(* IEC 61131-3 sources: Codesys_IAP/Demo/PLC1/Magazijn Overzetter Simulatie Structured Text 2V1_tekst/Simulatie, 5 files *)

(* ---- MagazijnDUT.st ---- *)
(*#### DECLARATIE ####*)
{attribute 'qualified_only'}
{attribute 'strict'}
TYPE MagazijnDUT :
(
	INGETROKKEN, INTREKKEN, UITGESTOTEN, UITSTOTEN, LEEG
);
END_TYPE

(* ---- OverzetterDUT.st ---- *)
(*#### DECLARATIE ####*)
{attribute 'qualified_only'}
{attribute 'strict'}
TYPE OverzetterDUT :
(
	INHETMIDDEN, NAARRECHTS, ISRECHTS, NAARLINKS, ISLINKS, GEVALLEN
);
END_TYPE

(* ---- SIM.st ---- *)
(*#### DECLARATIE ####*)
{attribute 'qualified_only'}
VAR_GLOBAL
	// Rotatie van de overzetter
	Vx_OvzRotate: INT := 0;
	// Visualisatie invisible blok
	Vx_OvzBlokLinks: BOOL := FALSE;
	// Visualisatie invisible blok
	Vx_OvzBlokOverzetter: BOOL := FALSE;
	// Visualisatie invisible blok
	Vx_OvzBlokRechts: BOOL := FALSE;
	// Visualisatie invisible blok
	Vx_OvzBlokGevallen: BOOL := FALSE;
	// Magazijn opnieuw vullen (simulatie)
	Ix_MagazijnVullen 	: BOOL;
	// Simulatie visualisatie
	Vw_Rotate45: INT := 45;
	// Visualisatie X positie van de uitstoter
	Vw_MagUitstoterBekerX: INT := 30;
	// Visualisatie invisible blok uitgestoten
	Vx_MagBlokUit: BOOL := TRUE;
	// Visualisatie invisible blok 1
	Vx_MagBlok1: BOOL := TRUE;
	// Visualisatie invisible blok 2
	Vx_MagBlok2: BOOL := TRUE;
	// Visualisatie invisible blok 3
	Vx_MagBlok3: BOOL := TRUE;
	// Visualisatie invisible blok 4
	Vx_MagBlok4: BOOL := TRUE;
	// Visualisatie invisible blokken
	Vx_MagBlok: ARRAY[1..8] OF BOOL;
	// Aantal blokken in het magazijn
	Vw_MagBlokAantal: INT := 4;
	// Simulatie onthoudt dat een blok maar 1x wordt uitgestoten
	Vw_MagBlok1X: INT := 0;
	// Simulatie error. Inverse logica.
	Vx_MagLuchtDrukError: BOOL := TRUE;
	// Simulatie error. Inverse logica.
	Vx_MagIsInError: BOOL := TRUE;
	// Simulatie error. Inverse logica.
	Vx_MagIsUitError: BOOL := TRUE;
	// Simulatie error. Inverse logica.
	Vx_OvzLuchtDrukError: BOOL := TRUE;
	// Simulatie error. Inverse logica.
	Vx_OvzIsLinksError: BOOL := TRUE;
	// Simulatie error. Inverse logica.
	Vx_OvzIsRechtsError: BOOL := TRUE;
	// Simulatie error. Inverse logica.
	Vx_OvzVacuumError: BOOL := TRUE;
	// Kleur van de blokken in het magazijn (lege plek = grijs)
	Vw_MagKleur: ARRAY[1..8] OF DWORD;
	// Kleur van het uitgestoten blok
	Vw_MagKleurUit: DWORD;
	// Kleur van het blok op de overzetter
	Vw_OvzKleur: DWORD := 16#FFC0C0C0;
	// Kleur van het blok dat klaarligt bij de uitgang van het magazijn
	Vw_MagKleurAfgifte: DWORD := 16#FFC0C0C0;
	// Er ligt een uitgestoten beker klaar bij de uitgang van het magazijn (voor de overzetter)
	Vx_MagBlokKlaar: BOOL := FALSE;
	// Afgifteplaats: kleur van de laatst afgegeven beker
	Vw_AfgifteKleur: DWORD := 16#FFA9A9A9;
	// Afgifteplaats: visualisatie invisible beker (inverse logica)
	Vx_AfgifteBeker: BOOL := TRUE;
	// Afgifteplaats: aantal afgegeven bekers
	Vi_AfgifteTeller: INT := 0;
	// Afgifteplaats leegmaken en teller op 0 (simulatie)
	Ix_AfgifteLegen: BOOL;
END_VAR

(* ---- MagazijnSim.st ---- *)
(*#### DECLARATIE ####*)
PROGRAM MagazijnSim
VAR
	// Timer om uitstoten en intrekken te vertragen
	Fb_Pulse: BLINK;
	// Timer om intrekken te vertragen
	Fb_Trigger: F_TRIG;
	// Eerste keer om visualisatie te updaten
	Mx_FirstTime: BOOL := TRUE;
	// Afhandeling van het magazijn
	Me_MagState: MAGAZIJNDUT := MAGAZIJNDUT.INGETROKKEN;
	// Kleuren van de blokken in het magazijn, [1] = onderste (wordt als eerste uitgestoten)
	Mw_KleurRij: ARRAY[1..8] OF DWORD;
	// Hulpvariabelen voor het kiezen van een willekeurige kleur
	Mi_Indx: INT;
	Mu_Seed: UDINT := 1;
END_VAR
VAR CONSTANT
	// Metaal blank (zilver): metaal en reflecterend
	METAAL_BLANK: DWORD := 16#FFC0C0C0;
	// Metaal zwart (antraciet): metaal, niet reflecterend
	METAAL_ZWART: DWORD := 16#FF505050;
	// Kunststof rood: geen metaal, wel reflecterend
	KUNSTOF_ROOD: DWORD := 16#FFFF0000;
	// Kunststof zwart: geen metaal, niet reflecterend
	KUNSTOF_ZWART: DWORD := 16#FF000000;
	// Lege plek in het magazijn
	LEEG: DWORD := 16#FFA9A9A9;
END_VAR
(*#### IMPLEMENTATIE ####*)
//
// Common stuff.
//

IF (Mx_FirstTime) THEN
	SIM.Vw_MagBlokAantal := 8;
	SIM.Vx_MagBlokUit:= FALSE;

	// Vul het magazijn met blokken in willekeurige kleuren (materiaal + kleur).
	Mu_Seed := DINT_TO_UDINT(TIME_TO_DINT(TIME())) + Mu_Seed;
	FOR Mi_Indx := 1 TO 8 DO
		Mu_Seed := Mu_Seed * 1103515245 + 12345;
		CASE UDINT_TO_INT(SHR(Mu_Seed, 16) AND 3) OF
			0: Mw_KleurRij[Mi_Indx] := METAAL_BLANK;
			1: Mw_KleurRij[Mi_Indx] := METAAL_ZWART;
			2: Mw_KleurRij[Mi_Indx] := KUNSTOF_ROOD;
		ELSE
			Mw_KleurRij[Mi_Indx] := KUNSTOF_ZWART;
		END_CASE
	END_FOR
	Mx_FirstTime := FALSE;
END_IF

//
// Handle all pulse and trigger events.
//
Fb_Pulse(ENABLE:=TRUE,TIMELOW:=T#200MS, TIMEHIGH:=T#200MS);
Fb_Trigger(CLK:=Fb_Pulse.OUT);

//
// Only if no emergency active, start handling the simulation.
//
IF (SIM.Ix_MagazijnVullen) THEN
	Mx_FirstTime := TRUE;
	SIM.Ix_MagazijnVullen := FALSE;
	RETURN;
END_IF

//
// The pulse determines the speed of the cilinder to move in
// ore move out. The cilinder is only moved if the airpressure
// is available.
//
IF (Fb_Trigger.Q AND SIM.Vx_MagLuchtDrukError) THEN

	CASE Me_MagState OF
		MAGAZIJNDUT.INGETROKKEN:
			IF (SIM.Vx_MagBlokUit) THEN
				SIM.Vw_MagBlokAantal := SIM.Vw_MagBlokAantal - 1;
				// Het onderste blok ligt nu klaar voor de overzetter; de rest zakt een plek.
				SIM.Vw_MagKleurAfgifte := Mw_KleurRij[1];
				SIM.Vx_MagBlokKlaar := TRUE;
				FOR Mi_Indx := 1 TO 7 DO
					Mw_KleurRij[Mi_Indx] := Mw_KleurRij[Mi_Indx + 1];
				END_FOR
				Mw_KleurRij[8] := LEEG;
			END_IF

			SIM.Vw_MagUitstoterBekerX := 1;
			SIM.Vw_MagBlok1X    	  := SIM.Vw_MagUitstoterBekerX;
			SIM.Vx_MagBlokUit         := FALSE;

			IF (Qx_BekerUitstoten) THEN
				Me_MagState := MAGAZIJNDUT.UITSTOTEN;
			END_IF

		MAGAZIJNDUT.INTREKKEN:
			SIM.Vw_MagUitstoterBekerX := SIM.Vw_MagUitstoterBekerX - 30;

			IF (SIM.Vw_MagUitstoterBekerX < 0) THEN
				SIM.Vw_MagUitstoterBekerX := 0;
			END_IF

			IF (SIM.Vw_MagUitstoterBekerX = 0) THEN
				Me_MagState := MAGAZIJNDUT.INGETROKKEN;
			END_IF

			IF (Qx_BekerUitstoten) THEN
				Me_MagState := MAGAZIJNDUT.UITSTOTEN;
			END_IF

		MAGAZIJNDUT.UITGESTOTEN:
			SIM.Vx_MagBlokUit         := SIM.Vx_MagBlok1;

			IF (NOT Qx_BekerUitstoten) THEN
				Me_MagState := MAGAZIJNDUT.INTREKKEN;
			END_IF

		MAGAZIJNDUT.UITSTOTEN:
			SIM.Vw_MagUitstoterBekerX := SIM.Vw_MagUitstoterBekerX + 30;
			SIM.Vw_MagBlok1X    	  := SIM.Vw_MagUitstoterBekerX;

			IF (SIM.Vw_MagUitstoterBekerX > 70) THEN
				Me_MagState := MAGAZIJNDUT.UITGESTOTEN;
			END_IF

			IF (NOT Qx_BekerUitstoten) THEN
				Me_MagState := MAGAZIJNDUT.INTREKKEN;
			END_IF

	END_CASE

	GVL.Ix_UitstoterBekerIn  := (Me_MagState = MAGAZIJNDUT.INGETROKKEN) AND SIM.Vx_MagIsInError;
	GVL.Ix_UitstoterBekerUit := (Me_MagState = MAGAZIJNDUT.UITGESTOTEN) AND SIM.Vx_MagIsUitError;
	GVL.Ix_MagazijnLeeg 	 := (SIM.Vw_MagBlokAantal <= 0) AND (Ix_UitstoterBekerIn);

	SIM.Vx_MagBlok[8] := (SIM.Vw_MagBlokAantal >= 8);
	SIM.Vx_MagBlok[7] := (SIM.Vw_MagBlokAantal >= 7);
	SIM.Vx_MagBlok[6] := (SIM.Vw_MagBlokAantal >= 6);
	SIM.Vx_MagBlok[5] := (SIM.Vw_MagBlokAantal >= 5);
	SIM.Vx_MagBlok[4] := (SIM.Vw_MagBlokAantal >= 4);
	SIM.Vx_MagBlok[3] := (SIM.Vw_MagBlokAantal >= 3);
	SIM.Vx_MagBlok[2] := (SIM.Vw_MagBlokAantal >= 2);
	SIM.Vx_MagBlok[1] := (SIM.Vw_MagBlokAantal >= 1);

	// Kleur per plek voor de visualisatie
	FOR Mi_Indx := 1 TO 8 DO
		IF SIM.Vx_MagBlok[Mi_Indx] THEN
			SIM.Vw_MagKleur[Mi_Indx] := Mw_KleurRij[Mi_Indx];
		ELSE
			SIM.Vw_MagKleur[Mi_Indx] := LEEG;
		END_IF
	END_FOR
	IF SIM.Vx_MagBlokUit THEN
		SIM.Vw_MagKleurUit := Mw_KleurRij[1];
	ELSE
		SIM.Vw_MagKleurUit := LEEG;
	END_IF

END_IF

(* ---- OverzetterSim.st ---- *)
(*#### DECLARATIE ####*)
PROGRAM OverzetterSim
VAR
	// Timer om overzetten te vertragen
	Fb_Pulse: BLINK;
	// Timer om overzetten te vertragen
	Fb_Trigger: F_TRIG;
	// Eerste keer om visualisatie te updaten
	Mx_FirstTime: BOOL := TRUE;
	// Afhandeling van de overzetter
	Me_OvzState: OverzetterDUT := OVERZETTERDUT.INHETMIDDEN;
	// Afhandeling van het blokje
	Me_BlokState: OverzetterDUT := OVERZETTERDUT.INHETMIDDEN;
	// Duurt even voor het vacuum aanwezig is
	Mi_VacuumCntr: INT := 0;
	// De overzetter heeft echt een beker vast (FALSE = leeg opgepakt, er lag niets klaar)
	Mx_MetBeker: BOOL := FALSE;
END_VAR
VAR CONSTANT

	// Inverse logica
	INVISABLE: BOOL := TRUE;
	// Inverse logica
	VISABLE: BOOL := FALSE;

END_VAR
(*#### IMPLEMENTATIE ####*)
// Initialisatie.

//
// Afgifteplaats leegmaken (knop in de visualisatie).
//
IF (SIM.Ix_AfgifteLegen) THEN
	SIM.Vi_AfgifteTeller := 0;
	SIM.Vx_AfgifteBeker  := INVISABLE;
	SIM.Vw_AfgifteKleur  := 16#FFA9A9A9;
	SIM.Ix_AfgifteLegen  := FALSE;
END_IF

IF (Mx_FirstTime) THEN
	Me_OvzState := OVERZETTERDUT.INHETMIDDEN;
	Me_BlokState := OVERZETTERDUT.ISLINKS;

	Mi_VacuumCntr := 0;
	Mx_MetBeker := FALSE;
	SIM.Vx_OvzRotate := 0;
	Mx_FirstTime := FALSE;
END_IF

//
// Afhandelen van de pulse events. Hierdoor loopt de simulatie los van de
// TASK tijd.
//
Fb_Pulse(ENABLE:=TRUE,TIMELOW:=T#100MS, TIMEHIGH:=T#100MS);
Fb_Trigger(CLK:=Fb_Pulse.OUT);

//
// Only if no emergency active, start handling the simulation.
//
IF (GVL.Ix_Noodstop) THEN
	Mx_FirstTime := TRUE;
	RETURN;
END_IF

//
// The pulse determines the speed of the cilinder to move in
// ore move out. The cilinder is only moved if the airpressure
// is available.
//
IF (Fb_Trigger.Q AND SIM.Vx_OvzLuchtDrukError) THEN

	//
	// De status van de arm wordt los afgehandeld van het blokje. De beweging
	// van de arm staat hier namelijk helemaal los van.
	//

	CASE Me_OvzState OF

		OVERZETTERDUT.INHETMIDDEN:
			//
			// De arm is in beweging naar links of naar rechts.
			// Indien de arm in de uiterste positie is wordt er van
			// state gewisseld. Aangezien de arm in beweging is staan
			// de eindschakelaars uit.
			//

			IF (GVL.Qx_OverzetterLinks) THEN
				IF (SIM.Vx_OvzRotate > -90) THEN
					GVL.Ix_OverzetterIsLinks := FALSE;
					GVL.Ix_OverzetterIsRechts := FALSE;
					SIM.Vx_OvzRotate := SIM.Vx_OvzRotate - 10;
				ELSE
					Me_OvzState := OVERZETTERDUT.ISLINKS;
				END_IF

			END_IF

			IF (GVL.Qx_OverzetterRechts) THEN
				IF (SIM.Vx_OvzRotate < 90) THEN
					GVL.Ix_OverzetterIsLinks := FALSE;
					GVL.Ix_OverzetterIsRechts := FALSE;
					SIM.Vx_OvzRotate := SIM.Vx_OvzRotate + 10;
				ELSE
					Me_OvzState := OVERZETTERDUT.ISRECHTS;
				END_IF
			END_IF

		OVERZETTERDUT.ISLINKS:
		    //
			// Arm staat in een uiterste stand. Eindschakelaar is ingeschakeld.
			// Zodra de arm weer wordt bewogen verandert de state.
			//

			GVL.Ix_OverzetterIsLinks := TRUE AND SIM.Vx_OvzIsLinksError;

			IF (GVL.Qx_OverzetterRechts AND NOT GVL.Qx_OverzetterLinks) THEN
				GVL.Ix_OverzetterIsLinks := FALSE;
				Me_OvzState := OVERZETTERDUT.INHETMIDDEN;
			END_IF

		OVERZETTERDUT.ISRECHTS:
		    //
			// Arm staat in een uiterste stand. Eindschakelaar is ingeschakeld.
			// Zodra de arm weer wordt bewogen verandert de state.
			//

			GVL.Ix_OverzetterIsRechts := TRUE AND SIM.Vx_OvzIsRechtsError;

			IF (GVL.Qx_OverzetterLinks AND NOT GVL.Qx_OverzetterRechts) THEN
				GVL.Ix_OverzetterIsRechts := FALSE;
				Me_OvzState := OVERZETTERDUT.INHETMIDDEN;
			END_IF

		END_CASE

	END_IF

	//
	// De status van het blokje hangt af van een aantal stuursignalen zoals waar
	// de arm zich bevindt, of er vacuum is en of er een beker lossen wordt gegeven.
	//

	CASE Me_BlokState OF
		OVERZETTERDUT.ISLINKS:
			//
			// Als de arm links is moet er eerst een vacuum opgebouwd worden alvorens het blokje
			// opgepakt kan worden. Daarna verandert de state. Er ligt alleen een blokje links
			// als het magazijn er een heeft uitgestoten (SIM.Vx_MagBlokKlaar).
			//

			SIM.Vx_OvzBlokGevallen 	 := INVISABLE;
			SIM.Vx_OvzBlokLinks 	 := NOT SIM.Vx_MagBlokKlaar;
			SIM.Vx_OvzBlokOverzetter := INVISABLE;
			SIM.Vx_OvzBlokRechts 	 := INVISABLE;

			IF (GVL.Qx_VacuumAan AND SIM.Vx_OvzVacuumError AND GVL.Ix_OverzetterIsLinks) AND (NOT GVL.Qx_BekerLossen) THEN
				Mi_VacuumCntr := Mi_VacuumCntr + 1;
			END_IF

			IF (NOT GVL.Qx_VacuumAan AND SIM.Vx_OvzVacuumError) THEN
				Mi_VacuumCntr := 0;
			END_IF

			GVL.Ix_VacuumAanwezig := (Mi_VacuumCntr > 50);

			IF  ( GVL.Ix_VacuumAanwezig AND (Me_OvzState = OVERZETTERDUT.INHETMIDDEN)) THEN
				// Het blok wordt opgepakt en krijgt de kleur van het blok uit het magazijn.
				// Lag er geen blok klaar, dan beweegt de arm leeg (en komt er niets op de afgifteplaats).
				Mx_MetBeker := SIM.Vx_MagBlokKlaar;
				SIM.Vx_MagBlokKlaar := FALSE;
				SIM.Vw_OvzKleur := SIM.Vw_MagKleurAfgifte;
				Me_BlokState := OVERZETTERDUT.INHETMIDDEN;
			END_IF

		OVERZETTERDUT.INHETMIDDEN:
			//
			// Het blokje is in beweging zolang er vacuum is. Als er geen vacuum meer is
			// valt het blokje... Indien de arm helemaal rechts is kan het blokje gelost
			// worden op de afgifteplaats. Dit moet met een Bekerlossen ondanks het feit dat er
			// geen vacuum meer is....
			//

			SIM.Vx_OvzBlokGevallen 	 := INVISABLE;
			SIM.Vx_OvzBlokLinks 	 := NOT SIM.Vx_MagBlokKlaar;
			SIM.Vx_OvzBlokOverzetter := NOT Mx_MetBeker;
			SIM.Vx_OvzBlokRechts 	 := INVISABLE;

		 	IF (GVL.Ix_OverzetterIsRechts) AND (NOT GVL.Qx_VacuumAan) AND (GVL.Qx_BekerLossen) THEN
				GVL.Ix_VacuumAanwezig := FALSE;
				IF Mx_MetBeker THEN
					// Beker komt op de afgifteplaats: zelfde kleur, teller omhoog.
					SIM.Vw_AfgifteKleur  := SIM.Vw_OvzKleur;
					SIM.Vx_AfgifteBeker  := VISABLE;
					SIM.Vi_AfgifteTeller := SIM.Vi_AfgifteTeller + 1;
				END_IF
				Me_BlokState := OVERZETTERDUT.ISRECHTS;
				RETURN;
			END_IF

			IF (NOT GVL.Ix_OverzetterIsRechts) AND (NOT GVL.Ix_OverzetterIsLinks) AND(NOT GVL.Qx_VacuumAan) THEN
				GVL.Ix_VacuumAanwezig := FALSE;
				Me_BlokState := OVERZETTERDUT.GEVALLEN;
			END_IF

		OVERZETTERDUT.ISRECHTS:
		    //
			// Blokje is gelost op de afgifteplaats. Nu is het wachten tot de overzetter terug naar links wordt gestuurd.
			//

			SIM.Vx_OvzBlokGevallen 	 := INVISABLE;
			SIM.Vx_OvzBlokLinks 	 := NOT SIM.Vx_MagBlokKlaar;
			SIM.Vx_OvzBlokOverzetter := INVISABLE;
			SIM.Vx_OvzBlokRechts 	 := INVISABLE;

			IF (NOT GVL.Ix_OverzetterIsRechts) THEN
				Mx_MetBeker := FALSE;
				Me_BlokState := OVERZETTERDUT.ISLINKS;
			END_IF

		OVERZETTERDUT.GEVALLEN:
			//
			// Blokje is gevallen..... Situatie herstelt zich zodra de arm helemaal links staat.
			//

			SIM.Vx_OvzBlokGevallen 	 := NOT Mx_MetBeker;
			SIM.Vx_OvzBlokLinks 	 := NOT SIM.Vx_MagBlokKlaar;
			SIM.Vx_OvzBlokOverzetter := INVISABLE;
			SIM.Vx_OvzBlokRechts 	 := INVISABLE;

			IF (GVL.Ix_OverzetterIsLinks) THEN
				Mx_MetBeker := FALSE;
				Me_BlokState := OVERZETTERDUT.ISLINKS;
			END_IF
	END_CASE
